ABB RAPID module: GoHome.mod

%%%
  VERSION:1
  LANGUAGE:ENGLISH
%%%
MODULE MOD_GoHome

    ! -------------------------------
    ! Define customized variables here
    ! ...

	! Tool variables:
	PERS tooldata SuctionCup := [TRUE,[[-94.709,0.000,259.352],[0.00000000,0.00000000,0.00000000,1.00000000]],[1,[0,0,20],[1,0,0,0],0,0,0.005]];

	! Reference variables:
	PERS wobjdata World := [FALSE, TRUE, "", [[0,0,0],[1,0,0,0]],[[390.000,0.000,0.000],[1.00000000,0.00000000,0.00000000,0.00000000]]];

	PROC Main()
		ConfJ \On;
		ConfL \Off;
		! Program generated by VerticalBot Studio for ABB IRB 1200-5/0.9 on 25/10/2026 12:00:00
		! Using nominal kinematics.
		MoveAbsJ [[0.000000,0.000000,-20.000000,0.000000,30.170000,0.000000],[9E+09,9E+09,9E+09,9E+09,9E+09,9E+09]],v500,z1,SuctionCup \WObj:=World;
	ENDPROC

ENDMODULE
